{region 'Documentation'}
(*!
<summary>Observes reservation state at request entry on a real minimal Test Case.</summary>
<description>
Inherits the normal lifecycle and one real Assertion from SuiteIntegrationChild.
Request overrides only count and observe before delegating to the production method.
No reservation result, state, readiness or scheduling decision is simulated.
ClearRequestTrace clears evidence only, before the isolated scenario begins.
</description>
*)
{endregion}
FUNCTION_BLOCK ReservationChildProbe EXTENDS SuiteIntegrationChild
VAR
    FResetRequestCount : UINT;
    FStartRequestCount : UINT;
    FRequestsReserved : BOOL := TRUE;
END_VAR
VAR CONSTANT
    ExecutionBudget : UINT := 11;
END_VAR

SUPER^();

{region 'Documentation'}
(*!
<summary>Clears observations without changing production lifecycle state.</summary>
*)
{endregion}
METHOD PUBLIC ClearRequestTrace
FResetRequestCount := 0;
FStartRequestCount := 0;
FRequestsReserved := TRUE;
END_METHOD

{region 'Documentation'}
(*!
<summary>Observes the held Reset budget before delegating the request.</summary>
*)
{endregion}
METHOD PUBLIC RequestReset
FResetRequestCount := FResetRequestCount + 1;
FRequestsReserved := FRequestsReserved
    AND (ReservedEntryCount = GVL_Constants.TestCaseResetEventCount)
    AND (EventPublisher.ReservedEntryCount >= ReservedEntryCount);
SUPER^.RequestReset();
END_METHOD

{region 'Documentation'}
(*!
<summary>Retained request-entry observation for the isolated scenario.</summary>
*)
{endregion}
{attribute 'monitoring' := 'call'}
PROPERTY PUBLIC RequestsReserved : BOOL //! Retained request-entry observation for the isolated scenario.
GET
RequestsReserved := FRequestsReserved;
END_GET
END_PROPERTY

{region 'Documentation'}
(*!
<summary>Observes the complete single-Assertion execution budget before delegating.</summary>
*)
{endregion}
METHOD PUBLIC RequestStart
FStartRequestCount := FStartRequestCount + 1;
FRequestsReserved := FRequestsReserved
    AND (ReservedEntryCount = ExecutionBudget)
    AND (EventPublisher.ReservedEntryCount >= ReservedEntryCount);
SUPER^.RequestStart();
END_METHOD

{region 'Documentation'}
(*!
<summary>Retained request-entry observation for the isolated scenario.</summary>
*)
{endregion}
{attribute 'monitoring' := 'call'}
PROPERTY PUBLIC ResetRequestCount : UINT //! Retained request-entry observation for the isolated scenario.
GET
ResetRequestCount := FResetRequestCount;
END_GET
END_PROPERTY

{region 'Documentation'}
(*!
<summary>Retained request-entry observation for the isolated scenario.</summary>
*)
{endregion}
{attribute 'monitoring' := 'call'}
PROPERTY PUBLIC StartRequestCount : UINT //! Retained request-entry observation for the isolated scenario.
GET
StartRequestCount := FStartRequestCount;
END_GET
END_PROPERTY

END_FUNCTION_BLOCK

(* stored: Version 1.1.0.1
   POU ReservationChildProbe: Id {6f70b8ac-9379-429f-acf4-02d8a19de581}, SpecialFunc None
   Method ClearRequestTrace: Id {39159cf0-73f1-40ab-9808-95bb76672376}
   Method RequestReset: Id {7a6c365c-fff7-43b2-bf04-ba79acfcbd27}
   Property RequestsReserved: Id {3d2bc57a-0b86-4658-a51e-92f83f208a74}
   Get Get: Id {073d4ed2-98ec-449d-aa7f-6a4b895abdf1}
   Method RequestStart: Id {ecaf3563-c763-4286-a91b-5d0673c5062c}
   Property ResetRequestCount: Id {2c364994-fc23-4618-a083-e7de72548e39}
   Get Get: Id {66e0ffb7-eb40-4b9d-86e6-2860ca64a087}
   Property StartRequestCount: Id {8c1e8aa9-e3c9-409a-aa40-d1dfb4b64757}
   Get Get: Id {a38d8481-cdc5-4eb5-9968-907107e04474} *)
